(* IEC 61131-3 sources: kns-pump-station/tests/POUs/Station/FB_Ats_Test, 15 files *)

(* ---- AtsClearsWhenPumpAvailableAgain.method.decl.st ---- *)
// 04 §9.1, PMI-12 шаг 3: снятый АВР насос освобождается, когда снова доступен (сброшен, в Auto); KNS1.ATS
// снимается
METHOD PRIVATE AtsClearsWhenPumpAvailableAgain
VAR
    fbDut   : FB_Ats;                          // ФБ под тестом
    fbTime  : PL.FB_FakeTime;                  // подменное время, старт 1 ч
    stCfg   : ST_StationCfg;                   // уставки по умолчанию (uiDutyMax = 2)
    afbPump : ARRAY[1..3] OF FB_FakeMotorVfd;  // подменные насосы: доступны, Auto
    fbSink  : FB_FakeEventSink;                // подменный журнал
END_VAR

(* ---- EventNamesReplacementPump.method.decl.st ---- *)
// 04 §16, PMI-12: событие 101006 с номером насоса, получившего новый запрос в окне STN_ATS_WINDOW; замена позже
// окна — без события
METHOD PRIVATE EventNamesReplacementPump
VAR
    fbDut   : FB_Ats;                          // ФБ под тестом
    fbTime  : PL.FB_FakeTime;                  // подменное время, старт 1 ч
    stCfg   : ST_StationCfg;                   // уставки по умолчанию (uiDutyMax = 2)
    afbPump : ARRAY[1..3] OF FB_FakeMotorVfd;  // подменные насосы: доступны, Auto
    fbSink  : FB_FakeEventSink;                // подменный журнал
    fbDut2  : FB_Ats;                          // второй экземпляр: замены нет
    uiStep  : UINT;                            // шаг 100 мс
END_VAR

(* ---- EventNamesReplacementPump.method.impl.st ---- *)
coUnit.TEST('Ats_EventNamesReplacementPump_A9_A16_PMI12');

fbDut.aitfPump[1] := afbPump[1];
fbDut.aitfPump[2] := afbPump[2];
fbDut.aitfPump[3] := afbPump[3];
fbDut.itfEvents := fbSink;
fbDut.xEnable := TRUE;
fbDut.uiAvailable := 3;

fbDut.axRun[1] := TRUE;
fbDut(itfTime := fbTime, stCfg := stCfg);
fbTime.Advance(tStep := T#100MS);

afbPump[1].xFault := TRUE;
fbDut.axRun[1] := FALSE;
fbDut(itfTime := fbTime, stCfg := stCfg);
AssertFalse(Condition := fbSink.Has(eFind := E_StationEvent.AtsPumpIn), Message := 'no replacement yet');
fbTime.Advance(tStep := T#1S);
fbDut.axRun[3] := TRUE;
fbDut(itfTime := fbTime, stCfg := stCfg);
AssertEquals_REAL(Expected := 3.0, Actual := fbSink.ValueOf(eFind := E_StationEvent.AtsPumpIn), Delta := 0.0,
                  Message := 'event 101006 names pump 3');
fbSink.Clear();
fbDut2.aitfPump[1] := afbPump[2];
fbDut2.itfEvents := fbSink;
fbDut2.xEnable := TRUE;
fbDut2.axRun[1] := TRUE;
fbDut2(itfTime := fbTime, stCfg := stCfg);
afbPump[2].xFault := TRUE;
fbDut2.axRun[1] := FALSE;
fbDut2(itfTime := fbTime, stCfg := stCfg);
FOR uiStep := 1 TO 101 DO
    fbTime.Advance(tStep := T#100MS);
    fbDut2(itfTime := fbTime, stCfg := stCfg);
END_FOR
fbDut2.axRun[2] := TRUE;
fbDut2(itfTime := fbTime, stCfg := stCfg);
AssertFalse(Condition := fbSink.Has(eFind := E_StationEvent.AtsPumpIn),
            Message := 'request after the window: no event');

coUnit.TEST_FINISHED();

(* ---- ForeignRunningCountsAgainstLack.method.decl.st ---- *)
// 04 §5.1, PMI-31: сторонний работающий насос откачивает — учитывается против нехватки
METHOD PRIVATE ForeignRunningCountsAgainstLack
VAR
    fbDut   : FB_Ats;                          // ФБ под тестом
    fbTime  : PL.FB_FakeTime;                  // подменное время, старт 1 ч
    stCfg   : ST_StationCfg;                   // уставки по умолчанию (uiDutyMax = 2)
    afbPump : ARRAY[1..3] OF FB_FakeMotorVfd;  // подменные насосы: доступны, Auto
    fbSink  : FB_FakeEventSink;                // подменный журнал
END_VAR

(* ---- LackWhenRequiredExceedsAvailable.method.decl.st ---- *)
// 04 §9.1, PMI-17: требуется больше насосов, чем доступно и работает стороннее, — условие KNS1.LACK
METHOD PRIVATE LackWhenRequiredExceedsAvailable
VAR
    fbDut   : FB_Ats;                          // ФБ под тестом
    fbTime  : PL.FB_FakeTime;                  // подменное время, старт 1 ч
    stCfg   : ST_StationCfg;                   // уставки по умолчанию (uiDutyMax = 2)
    afbPump : ARRAY[1..3] OF FB_FakeMotorVfd;  // подменные насосы: доступны, Auto
    fbSink  : FB_FakeEventSink;                // подменный журнал
END_VAR

(* ---- ModeChangeIsNotAts.method.decl.st ---- *)
// 04 §9.1, PMI-31: перевод запрошенного насоса в Local оператором — не АВР
METHOD PRIVATE ModeChangeIsNotAts
VAR
    fbDut   : FB_Ats;                          // ФБ под тестом
    fbTime  : PL.FB_FakeTime;                  // подменное время, старт 1 ч
    stCfg   : ST_StationCfg;                   // уставки по умолчанию (uiDutyMax = 2)
    afbPump : ARRAY[1..3] OF FB_FakeMotorVfd;  // подменные насосы: доступны, Auto
    fbSink  : FB_FakeEventSink;                // подменный журнал
END_VAR

(* ---- NoReserveUsesEffectiveDuty.method.decl.st ---- *)
// 04 §5.1, §6, §7.2, §15, PMI-32: в обычном режиме работает не больше MIN(uiDutyMax, STN_DUTY_MAX) насосов
// (ступенчатое и ПИД — до двух). При допустимом uiDutyMax = 3 три доступных насоса — это два рабочих и резерв:
// условие KNS1.NORES ложно (иначе постоянная High-тревога при исправной станции)
METHOD PRIVATE NoReserveUsesEffectiveDuty
VAR
    fbDut   : FB_Ats;                          // ФБ под тестом
    fbTime  : PL.FB_FakeTime;                  // подменное время, старт 1 ч
    stCfg   : ST_StationCfg;                   // уставки по умолчанию, uiDutyMax = 3
    afbPump : ARRAY[1..3] OF FB_FakeMotorVfd;  // подменные насосы: доступны, Auto
    fbSink  : FB_FakeEventSink;                // подменный журнал
END_VAR

(* ---- NoReserveWhenOnePumpUnavailable.method.decl.st ---- *)
// 04 §15, PMI-32: доступно меньше uiDutyMax + 1 — условие KNS1.NORES
METHOD PRIVATE NoReserveWhenOnePumpUnavailable
VAR
    fbDut   : FB_Ats;                          // ФБ под тестом
    fbTime  : PL.FB_FakeTime;                  // подменное время, старт 1 ч
    stCfg   : ST_StationCfg;                   // уставки по умолчанию (uiDutyMax = 2)
    afbPump : ARRAY[1..3] OF FB_FakeMotorVfd;  // подменные насосы: доступны, Auto
    fbSink  : FB_FakeEventSink;                // подменный журнал
END_VAR

(* ---- PowerLossIsNotAts.method.decl.st ---- *)
// 04 §9.1, PMI-33: пропадание напряжения (насос недоступен без отказа) — не АВР
METHOD PRIVATE PowerLossIsNotAts
VAR
    fbDut   : FB_Ats;                          // ФБ под тестом
    fbTime  : PL.FB_FakeTime;                  // подменное время, старт 1 ч
    stCfg   : ST_StationCfg;                   // уставки по умолчанию (uiDutyMax = 2)
    afbPump : ARRAY[1..3] OF FB_FakeMotorVfd;  // подменные насосы: доступны, Auto
    fbSink  : FB_FakeEventSink;                // подменный журнал
END_VAR

(* ---- RequestedPumpFaultRaisesAts.method.decl.st ---- *)
// 04 §9.1, PMI-12, PMI-13: отказ насоса, запрошенного в прошлом цикле, — АВР: насос снят, KNS1.ATS, счётчик АВР
METHOD PRIVATE RequestedPumpFaultRaisesAts
VAR
    fbDut   : FB_Ats;                          // ФБ под тестом
    fbTime  : PL.FB_FakeTime;                  // подменное время, старт 1 ч
    stCfg   : ST_StationCfg;                   // уставки по умолчанию (uiDutyMax = 2)
    afbPump : ARRAY[1..3] OF FB_FakeMotorVfd;  // подменные насосы: доступны, Auto
    fbSink  : FB_FakeEventSink;                // подменный журнал
END_VAR

(* ---- TimeBackwardsWindowRestarts.method.decl.st ---- *)
// Время назад — окно STN_ATS_WINDOW отсчитывается заново, замена в окне называется в событии 101006
METHOD PRIVATE TimeBackwardsWindowRestarts
VAR
    fbDut   : FB_Ats;                          // ФБ под тестом
    fbTime  : PL.FB_FakeTime;                  // подменное время, старт 1 ч
    stCfg   : ST_StationCfg;                   // уставки по умолчанию (uiDutyMax = 2)
    afbPump : ARRAY[1..3] OF FB_FakeMotorVfd;  // подменные насосы: доступны, Auto
    fbSink  : FB_FakeEventSink;                // подменный журнал
    uiStep  : UINT;                            // шаг 100 мс
END_VAR

(* ---- TimeBackwardsWindowRestarts.method.impl.st ---- *)
coUnit.TEST('Ats_TimeBackwardsWindowRestarts_A9');

fbDut.aitfPump[1] := afbPump[1];
fbDut.aitfPump[2] := afbPump[2];
fbDut.aitfPump[3] := afbPump[3];
fbDut.itfEvents := fbSink;
fbDut.xEnable := TRUE;
fbDut.uiAvailable := 3;

fbDut.axRun[1] := TRUE;
fbDut(itfTime := fbTime, stCfg := stCfg);
fbTime.Advance(tStep := T#100MS);

afbPump[1].xFault := TRUE;
fbDut.axRun[1] := FALSE;
fbDut(itfTime := fbTime, stCfg := stCfg);
fbTime.SetNow(ltValue := LTIME#59M);
FOR uiStep := 1 TO 95 DO
    fbTime.Advance(tStep := T#100MS);
    fbDut(itfTime := fbTime, stCfg := stCfg);
END_FOR
fbDut.axRun[2] := TRUE;
fbDut(itfTime := fbTime, stCfg := stCfg);
AssertEquals_REAL(Expected := 2.0, Actual := fbSink.ValueOf(eFind := E_StationEvent.AtsPumpIn), Delta := 0.0,
                  Message := 'replacement inside restarted window');

coUnit.TEST_FINISHED();

(* ---- TripEventNamesReplacementNotTrippedPump.method.decl.st ---- *)
// 04 §9.1, §16, PMI-15, PMI-16: блокировка станции (недогрузка, перегрев) — в цикле отказа насос ещё доступен и
// запрошен (FB_PumpRotation снимет запрос со следующего цикла). Событие 101006 называет замену, а не сам снятый АВР
// насос
METHOD PRIVATE TripEventNamesReplacementNotTrippedPump
VAR
    fbDut   : FB_Ats;                          // ФБ под тестом
    fbTime  : PL.FB_FakeTime;                  // подменное время, старт 1 ч
    stCfg   : ST_StationCfg;                   // уставки по умолчанию (uiDutyMax = 2)
    afbPump : ARRAY[1..3] OF FB_FakeMotorVfd;  // подменные насосы: доступны, Auto
    fbSink  : FB_FakeEventSink;                // подменный журнал
END_VAR

(* ---- UnderloadTripIsAts.method.decl.st ---- *)
// 04 §9.1, PMI-15: фиксация недогрузки станцией (axTrip) у запрошенного насоса — АВР, даже пока устройство ещё
// доступно; снят, пока фиксация не сброшена
METHOD PRIVATE UnderloadTripIsAts
VAR
    fbDut   : FB_Ats;                          // ФБ под тестом
    fbTime  : PL.FB_FakeTime;                  // подменное время, старт 1 ч
    stCfg   : ST_StationCfg;                   // уставки по умолчанию (uiDutyMax = 2)
    afbPump : ARRAY[1..3] OF FB_FakeMotorVfd;  // подменные насосы: доступны, Auto
    fbSink  : FB_FakeEventSink;                // подменный журнал
END_VAR

(* ---- UnrequestedOrManualFaultIsNotAts.method.decl.st ---- *)
// 04 §9.1, PMI-14: отказ незапрошенного насоса и отказ в «Ручном» станции — не АВР
METHOD PRIVATE UnrequestedOrManualFaultIsNotAts
VAR
    fbDut   : FB_Ats;                          // ФБ под тестом
    fbTime  : PL.FB_FakeTime;                  // подменное время, старт 1 ч
    stCfg   : ST_StationCfg;                   // уставки по умолчанию (uiDutyMax = 2)
    afbPump : ARRAY[1..3] OF FB_FakeMotorVfd;  // подменные насосы: доступны, Auto
    fbSink  : FB_FakeEventSink;                // подменный журнал
END_VAR
